(* IEC 61131-3 sources: Lasal-MCP/examples/SampleSource/5_ClassInputOutputSolution/Stations/MachineControl/MachineControl/Class/OPModeConfigBase, 1 file *)

(* ---- OPModeConfigBase.st ---- *)
#define     NewInstCmd_GetAlarms                  100     // newinst command to get alarms of station (class AlarmSation + class OPModeComMaster)
// parameter 1: sAlarmList  : t_s_OPMode
// parameter 2: bdAlarmInfo : BDINT

(*!
<Class
	Name               = "OPModeConfigBase"
	Revision           = "1.3"
	RealtimeTask       = "false"
	CyclicTask         = "false"
	BackgroundTask     = "false"
	Sigmatek           = "true"
	OSInterface        = "false"
	HighPriority       = "false"
	Automatic          = "false"
	UpdateMode         = "Prescan"
	SharedCommandTable = "true"
	Objectsize         = "(410,120)"
	Comment            = "This class defines the configuration for the class OPModeBase.&#13;&#10;All the possible ways to change the operation mode are defined within this class.&#13;&#10;&#13;&#10;Derive this class to change the configuration for switching the operation modes.">
	<Channels>
		<Server Name="ClassSvr" Visualized="false" Initialize="false" WriteProtected="true" Retentive="false"/>
	</Channels>
	<RevDoku>
		<Owner Company="Sigmatek" Author="ObeChr"/>
		<Dokumentation Revision="1.3" Date="2018-04-17" Author="ObeChr" Company="Sigmatek" Description="Added functionality that it is possible to call Change-Methods until every Slave Object is READY"/>
		<Dokumentation Revision="1.2" Date="2017-01-30" Author="ObeChr" Company="Sigmatek" Description="Added new public types to class."/>
		<Dokumentation Revision="1.1" Date="2016-03-08" Author="ObeChr" Company="Sigmatek" Description="+) Added deactivated configurations to the methods GetChangeConfig(), GetModeConfig() to show the possibilties of the class.&#13;&#10;+) Deactivated all transition times.&#13;&#10;+) Improved comments of global methods and variables."/>
		<Dokumentation Revision="1.0" Date="2015-06-01" Author="ObeChr" Company="Sigmatek" Description="First Version of class for the configuration of the operationmodes."/>
	</RevDoku>
</Class>
*)
OPModeConfigBase : CLASS
	TYPE
	  t_bd_OPMode : BDINT  //! <Type Public="true" Name="t_bd_OPMode"/>
	  [
	    1 bOPModeInit,
	    2 bOPModeHoming,
	    3 bOPModeStop,
	    4 bOPModeSetup,
	    5 bOPModeManual,
	    6 bOPModeSemiAuto,
	    7 bOPModeAutomatic,
	    8 bOPModeError,
	  ];
#pragma pack(push, 1)
	  t_s_OPChange : STRUCT  //! <Type Public="true" Name="t_s_OPChange"/>
	    bOPModeInit : BINT  //! <Type Comment="This bit field defines the optional operating modes to which are changed from the operating mode Init." Name="t_s_OPChange.bOPModeInit"/>
	    [
	      1 bHoming,
	      2 bStop,
	      3 bSetup,
	      4 bManual,
	      5 bSemiAuto,
	      6 bAutomatic,
	      7 bError,
	    ];
	    bOPModeHoming : BINT  //! <Type Comment="This bit field defines the optional operating modes to which are changed from the operating mode Homing." Name="t_s_OPChange.bOPModeHoming"/>
	    [
	      1 bInit,
	      2 bStop,
	      3 bSetup,
	      4 bManual,
	      5 bSemiAuto,
	      6 bAutomatic,
	      7 bError,
	    ];
	    bOPModeStop : BINT  //! <Type Comment="This bit field defines the optional operating modes to which are changed from the operating mode Stop." Name="t_s_OPChange.bOPModeStop"/>
	    [
	      1 bInit,
	      2 bHoming,
	      3 bSetup,
	      4 bManual,
	      5 bSemiAuto,
	      6 bAutomatic,
	      7 bError,
	    ];
	    bOPModeSetup : BINT  //! <Type Comment="This bit field defines the optional operating modes to which are changed from the operating mode Setup." Name="t_s_OPChange.bOPModeSetup"/>
	    [
	      1 bInit,
	      2 bHoming,
	      3 bStop,
	      4 bManual,
	      5 bSemiAuto,
	      6 bAutomatic,
	      7 bError,
	    ];
	    bOPModeManual : BINT  //! <Type Comment="This bit field defines the optional operating modes to which are changed from the operating mode Manual." Name="t_s_OPChange.bOPModeManual"/>
	    [
	      1 bInit,
	      2 bHoming,
	      3 bStop,
	      4 bSetup,
	      5 bSemiAuto,
	      6 bAutomatic,
	      7 bError,
	    ];
	    bOPModeSemiAuto : BINT  //! <Type Comment="This bit field defines the optional operating modes to which are changed from the operating mode SemiAuto." Name="t_s_OPChange.bOPModeSemiAuto"/>
	    [
	      1 bInit,
	      2 bHoming,
	      3 bStop,
	      4 bSetup,
	      5 bManual,
	      6 bAutomatic,
	      7 bError,
	    ];
	    bOPModeAutomatic : BINT  //! <Type Comment="This bit field defines the optional operating modes to which are changed from the operating mode Automatic." Name="t_s_OPChange.bOPModeAutomatic"/>
	    [
	      1 bInit,
	      2 bHoming,
	      3 bStop,
	      4 bSetup,
	      5 bManual,
	      6 bSemiAuto,
	      7 bError,
	    ];
	    bOPModeError : BINT  //! <Type Comment="This bit field defines the optional operating modes to which are changed from the operating mode Error." Name="t_s_OPChange.bOPModeError"/>
	    [
	      1 bInit,
	      2 bHoming,
	      3 bStop,
	      4 bSetup,
	      5 bManual,
	      6 bSemiAuto,
	      7 bAutomatic,
	    ];
	  END_STRUCT;
#pragma pack(pop)
#pragma pack(push, 1)
	  t_s_OPChangeTime : STRUCT  //! <Type Public="true" Name="t_s_OPChangeTime"/>
	    sOPModeInit : STRUCT  //! <Type Comment="In this structure, the allowable changeover times [ms] are defined from OPMode_Init.&#13;&#10;" Name="t_s_OPChangeTime.sOPModeInit"/>
	      udChangeToHoming : UDINT;
	      udChangeToStop : UDINT;
	      udChangeToSetup : UDINT;
	      udChangeToManual : UDINT;
	      udChangeToSemiAuto : UDINT;
	      udChangeToAutomatic : UDINT;
	      udChangeToError : UDINT;
	    END_STRUCT;
	    sOPModeHoming : STRUCT  //! <Type Comment="In this structure, the allowable changeover times [ms] are defined from OPMode_Homing.&#13;&#10;" Name="t_s_OPChangeTime.sOPModeHoming"/>
	      udChangeToInit : UDINT;
	      udChangeToStop : UDINT;
	      udChangeToSetup : UDINT;
	      udChangeToManual : UDINT;
	      udChangeToSemiAuto : UDINT;
	      udChangeToAutomatic : UDINT;
	      udChangeToError : UDINT;
	    END_STRUCT;
	    sOPModeStop : STRUCT  //! <Type Comment="In this structure, the allowable changeover times [ms] are defined from OPMode_Stop.&#13;&#10;" Name="t_s_OPChangeTime.sOPModeStop"/>
	      udChangeToInit : UDINT;
	      udChangeToHoming : UDINT;
	      udChangeToSetup : UDINT;
	      udChangeToManual : UDINT;
	      udChangeToSemiAuto : UDINT;
	      udChangeToAutomatic : UDINT;
	      udChangeToError : UDINT;
	    END_STRUCT;
	    sOPModeSetup : STRUCT  //! <Type Comment="In this structure, the allowable changeover times [ms] are defined from OPMode_Setup.&#13;&#10;" Name="t_s_OPChangeTime.sOPModeSetup"/>
	      udChangeToInit : UDINT;
	      udChangeToHoming : UDINT;
	      udChangeToStop : UDINT;
	      udChangeToManual : UDINT;
	      udChangeToSemiAuto : UDINT;
	      udChangeToAutomatic : UDINT;
	      udChangeToError : UDINT;
	    END_STRUCT;
	    sOPModeManual : STRUCT  //! <Type Comment="In this structure, the allowable changeover times [ms] are defined from OPMode_Manual.&#13;&#10;" Name="t_s_OPChangeTime.sOPModeManual"/>
	      udChangeToInit : UDINT;
	      udChangeToHoming : UDINT;
	      udChangeToStop : UDINT;
	      udChangeToSetup : UDINT;
	      udChangeToSemiAuto : UDINT;
	      udChangeToAutomatic : UDINT;
	      udChangeToError : UDINT;
	    END_STRUCT;
	    sOPModeSemiAuto : STRUCT  //! <Type Comment="In this structure, the allowable changeover times [ms] are defined from OPMode_SemiAuto.&#13;&#10;" Name="t_s_OPChangeTime.sOPModeSemiAuto"/>
	      udChangeToInit : UDINT;
	      udChangeToHoming : UDINT;
	      udChangeToStop : UDINT;
	      udChangeToSetup : UDINT;
	      udChangeToManual : UDINT;
	      udChangeToAutomatic : UDINT;
	      udChangeToError : UDINT;
	    END_STRUCT;
	    sOPModeAutomatic : STRUCT  //! <Type Comment="In this structure, the allowable changeover times [ms] are defined from OPMode_Automatic.&#13;&#10;" Name="t_s_OPChangeTime.sOPModeAutomatic"/>
	      udChangeToInit : UDINT;
	      udChangeToHoming : UDINT;
	      udChangeToStop : UDINT;
	      udChangeToSetup : UDINT;
	      udChangeToManual : UDINT;
	      udChangeToSemiAuto : UDINT;
	      udChangeToError : UDINT;
	    END_STRUCT;
	    sOPModeError : STRUCT  //! <Type Comment="In this structure, the allowable changeover times [ms] are defined from OPMode_Error.&#13;&#10;" Name="t_s_OPChangeTime.sOPModeError"/>
	      udChangeToInit : UDINT;
	      udChangeToHoming : UDINT;
	      udChangeToStop : UDINT;
	      udChangeToSetup : UDINT;
	      udChangeToManual : UDINT;
	      udChangeToSemiAuto : UDINT;
	      udChangeToAutomatic : UDINT;
	    END_STRUCT;
	  END_STRUCT;
#pragma pack(pop)
	END_TYPE
  //Servers:
	ClassSvr 	: SvrChCmd_DINT;
  //Clients:
  //Variables:
		bdOPMode 	: t_bd_OPMode;			//! <Variable Comment="This variable defines the available operation modes." Name="bdOPMode"/>
		sOPChange 	: t_s_OPChange;			//! <Variable Comment="This variable defines the possible transitions between the operation modes." Name="sOPChange"/>
		sOPChangeTime 	: t_s_OPChangeTime;			//! <Variable Comment="This variable defines the timeouts for the transitions between the operation modes." Name="sOPChangeTime"/>
  //Functions:
				//! <Function Comment="This method is called by the &quot;OPModeBase&quot; class during the last Init cycle. The configuration of the class is thereby defined. By overwriting this method, the default configuration can be changed." Name="GetChangeConfig"/>
	FUNCTION VIRTUAL GLOBAL GetChangeConfig
		VAR_OUTPUT
			pConfig 	: ^t_s_OPChange;			//! <Variable Comment="Pointer to the changeover options of the operating mode (sOPModeChange variable)." Name="GetChangeConfig.pConfig"/>
		END_VAR;
				//! <Function Comment="This method is called by the &quot;OPModeBase&quot; class during the last Init cycle. Through this call, the configuration is read based on allowed changeover time of the operating modes. By overwriting this method, the default configuration can be changed." Name="GetChangeTime"/>
	FUNCTION VIRTUAL GLOBAL GetChangeTime
		VAR_OUTPUT
			pConfig 	: ^t_s_OPChangeTime;			//! <Variable Comment="Pointer to the timeouts when changing operating modes  (variable sOPChangeTime)." Name="GetChangeTime.pConfig"/>
		END_VAR;
				//! <Function Comment="This method is called by the &quot;AlarmBufferBase&quot; class when registering an alarm. The possible configuration of the alarm is checked. By overwriting this method, the default configuration can be changed." Name="GetModeConfig"/>
	FUNCTION VIRTUAL GLOBAL GetModeConfig
		VAR_OUTPUT
			pConfig 	: ^t_bd_OPMode;			//! <Variable Comment="Pointer to the available operating modes (variable bdOPMode)." Name="GetModeConfig.pConfig"/>
		END_VAR;
  //Tables:
	FUNCTION @STD
		VAR_OUTPUT
			ret_code	: CONFSTATES;
		END_VAR;
	FUNCTION GLOBAL TAB @CT_;
END_CLASS;

FUNCTION VIRTUAL GLOBAL OPModeConfigBase::GetChangeConfig
	VAR_OUTPUT
		pConfig 	: ^t_s_OPChange;
	END_VAR

  // this information is ued by the class OPModeBase
  // => only following transitions between the OPModes
  //    can be used

  // possibilities to leave OPMode_Init
  sOPChange.bOPModeInit.bHoming     := true;        // transition active
  sOPChange.bOPModeInit.bStop       := false;
  sOPChange.bOPModeInit.bSetup      := false;
  sOPChange.bOPModeInit.bManual     := false;
  sOPChange.bOPModeInit.bSemiAuto   := false;
  sOPChange.bOPModeInit.bAutomatic  := false;
  sOPChange.bOPModeInit.bError      := true;        // transition active

  // possibilities to leave OPMode_Homing
  sOPChange.bOPModeHoming.bInit       := false;
  sOPChange.bOPModeHoming.bStop       := false;
  sOPChange.bOPModeHoming.bSetup      := false;
  sOPChange.bOPModeHoming.bManual     := true;      // transition active
  sOPChange.bOPModeHoming.bSemiAuto   := false;
  sOPChange.bOPModeHoming.bAutomatic  := false;
  sOPChange.bOPModeHoming.bError      := true;      // transition active

  // possibilities to leave OPMode_Stop
  sOPChange.bOPModeStop.bInit       := false;
  sOPChange.bOPModeStop.bHoming     := false;
  sOPChange.bOPModeStop.bSetup      := false;
  sOPChange.bOPModeStop.bManual     := false;
  sOPChange.bOPModeStop.bSemiAuto   := false;
  sOPChange.bOPModeStop.bAutomatic  := false;
  sOPChange.bOPModeStop.bError      := false;

  // possibilities to leave OPMode_Setup
  sOPChange.bOPModeSetup.bInit      := false;
  sOPChange.bOPModeSetup.bHoming    := false;
  sOPChange.bOPModeSetup.bStop      := false;
  sOPChange.bOPModeSetup.bManual    := false;
  sOPChange.bOPModeSetup.bSemiAuto  := false;
  sOPChange.bOPModeSetup.bAutomatic := false;
  sOPChange.bOPModeSetup.bError     := false;

  // possibilities to leave OPMode_Manual
  sOPChange.bOPModeManual.bInit       := true;      // transition active
  sOPChange.bOPModeManual.bHoming     := true;      // transition active
  sOPChange.bOPModeManual.bStop       := false;
  sOPChange.bOPModeManual.bSetup      := false;
  sOPChange.bOPModeManual.bSemiAuto   := true;      // transition active
  sOPChange.bOPModeManual.bAutomatic  := true;      // transition active
  sOPChange.bOPModeManual.bError      := true;      // transition active

  // possibilities to leave OPMode_SemiAuto
  sOPChange.bOPModeSemiAuto.bInit       := false;
  sOPChange.bOPModeSemiAuto.bHoming     := false;
  sOPChange.bOPModeSemiAuto.bStop       := false;
  sOPChange.bOPModeSemiAuto.bSetup      := false;
  sOPChange.bOPModeSemiAuto.bManual     := true;    // transition active
  sOPChange.bOPModeSemiAuto.bAutomatic  := true;    // transition active
  sOPChange.bOPModeSemiAuto.bError      := true;    // transition active

  // possibilities to leave OPMode_Automatic
  sOPChange.bOPModeAutomatic.bInit      := false;
  sOPChange.bOPModeAutomatic.bHoming    := false;
  sOPChange.bOPModeAutomatic.bStop      := false;
  sOPChange.bOPModeAutomatic.bSetup     := false;
  sOPChange.bOPModeAutomatic.bManual    := true;    // transition active
  sOPChange.bOPModeAutomatic.bSemiAuto  := true;    // transition active
  sOPChange.bOPModeAutomatic.bError     := true;    // transition active

  // possibilities to leave OPMode_Error
  sOPChange.bOPModeError.bInit      := true;        // transition active
  sOPChange.bOPModeError.bHoming    := true;        // transition active
  sOPChange.bOPModeError.bStop      := false;
  sOPChange.bOPModeError.bSetup     := false;
  sOPChange.bOPModeError.bManual    := true;        // transition active
  sOPChange.bOPModeError.bSemiAuto  := false;
  sOPChange.bOPModeError.bAutomatic := false;

  // return pointer to configuration
  pConfig := #sOPChange;

END_FUNCTION

FUNCTION VIRTUAL GLOBAL OPModeConfigBase::GetModeConfig
	VAR_OUTPUT
		pConfig 	: ^t_bd_OPMode;
	END_VAR

  // this information is used by the class AlarmBuffer
  // => only following OPModes can be set at the alarm
  //    objects

  // available OPModes
  bdOPMode.bOPModeInit      := true;    // OPMode active
  bdOPMode.bOPModeHoming    := true;    // OPMode active
  bdOPMode.bOPModeStop      := false;
  bdOPMode.bOPModeSetup     := false;
  bdOPMode.bOPModeManual    := true;    // OPMode active
  bdOPMode.bOPModeSemiAuto  := true;    // OPMode active
  bdOPMode.bOPModeAutomatic := true;    // OPMode active
  bdOPMode.bOPModeError     := true;    // OPMode active

  // return configuration
  pConfig := #bdOPMode;

END_FUNCTION

FUNCTION VIRTUAL GLOBAL OPModeConfigBase::GetChangeTime
	VAR_OUTPUT
		pConfig 	: ^t_s_OPChangeTime;
	END_VAR

  // this information is ued by the class OPModeBase
  // => in case changing the opmode takes more than
  //    the selected time, an error occus.
  // 0: check of transitiontime is deactivated

  // timeouts to leave OPMode_Init
  sOPChangeTime.sOPModeInit.udChangeToHoming    := 0;
  sOPChangeTime.sOPModeInit.udChangeToStop      := 0;
  sOPChangeTime.sOPModeInit.udChangeToSetup     := 0;
  sOPChangeTime.sOPModeInit.udChangeToManual    := 0;
  sOPChangeTime.sOPModeInit.udChangeToSemiAuto  := 0;
  sOPChangeTime.sOPModeInit.udChangeToAutomatic := 0;
  sOPChangeTime.sOPModeInit.udChangeToError     := 0;

  // timeouts to leave OPMode_Homing
  sOPChangeTime.sOPModeHoming.udChangeToInit      := 0;
  sOPChangeTime.sOPModeHoming.udChangeToStop      := 0;
  sOPChangeTime.sOPModeHoming.udChangeToSetup     := 0;
  sOPChangeTime.sOPModeHoming.udChangeToManual    := 0;
  sOPChangeTime.sOPModeHoming.udChangeToSemiAuto  := 0;
  sOPChangeTime.sOPModeHoming.udChangeToAutomatic := 0;
  sOPChangeTime.sOPModeHoming.udChangeToError     := 0;

  // timeouts to leave OPMode_Stop
  sOPChangeTime.sOPModeStop.udChangeToInit      := 0;
  sOPChangeTime.sOPModeStop.udChangeToHoming    := 0;
  sOPChangeTime.sOPModeStop.udChangeToSetup     := 0;
  sOPChangeTime.sOPModeStop.udChangeToManual    := 0;
  sOPChangeTime.sOPModeStop.udChangeToSemiAuto  := 0;
  sOPChangeTime.sOPModeStop.udChangeToAutomatic := 0;
  sOPChangeTime.sOPModeStop.udChangeToError     := 0;

  // timeouts to leave OPMode_Setup
  sOPChangeTime.sOPModeSetup.udChangeToInit       := 0;
  sOPChangeTime.sOPModeSetup.udChangeToHoming     := 0;
  sOPChangeTime.sOPModeSetup.udChangeToStop       := 0;
  sOPChangeTime.sOPModeSetup.udChangeToManual     := 0;
  sOPChangeTime.sOPModeSetup.udChangeToSemiAuto   := 0;
  sOPChangeTime.sOPModeSetup.udChangeToAutomatic  := 0;
  sOPChangeTime.sOPModeSetup.udChangeToError      := 0;

  // timeouts to leave OPMode_Manual
  sOPChangeTime.sOPModeManual.udChangeToInit      := 0;
  sOPChangeTime.sOPModeManual.udChangeToHoming    := 0;
  sOPChangeTime.sOPModeManual.udChangeToStop      := 0;
  sOPChangeTime.sOPModeManual.udChangeToSetup     := 0;
  sOPChangeTime.sOPModeManual.udChangeToSemiAuto  := 0;
  sOPChangeTime.sOPModeManual.udChangeToAutomatic := 0;
  sOPChangeTime.sOPModeManual.udChangeToError     := 0;

  // timeouts to leave OPMode_SemiAuto
  sOPChangeTime.sOPModeSemiAuto.udChangeToInit      := 0;
  sOPChangeTime.sOPModeSemiAuto.udChangeToHoming    := 0;
  sOPChangeTime.sOPModeSemiAuto.udChangeToStop      := 0;
  sOPChangeTime.sOPModeSemiAuto.udChangeToSetup     := 0;
  sOPChangeTime.sOPModeSemiAuto.udChangeToManual    := 0;
  sOPChangeTime.sOPModeSemiAuto.udChangeToAutomatic := 0;
  sOPChangeTime.sOPModeSemiAuto.udChangeToError     := 0;

  // timeouts to leave OPMode_Automatic
  sOPChangeTime.sOPModeAutomatic.udChangeToInit     := 0;
  sOPChangeTime.sOPModeAutomatic.udChangeToHoming   := 0;
  sOPChangeTime.sOPModeAutomatic.udChangeToStop     := 0;
  sOPChangeTime.sOPModeAutomatic.udChangeToSetup    := 0;
  sOPChangeTime.sOPModeAutomatic.udChangeToManual   := 0;
  sOPChangeTime.sOPModeAutomatic.udChangeToSemiAuto := 0;
  sOPChangeTime.sOPModeAutomatic.udChangeToError    := 0;

  // timeouts to leave OPMode_Error
  sOPChangeTime.sOPModeError.udChangeToInit       := 0;
  sOPChangeTime.sOPModeError.udChangeToHoming     := 0;
  sOPChangeTime.sOPModeError.udChangeToStop       := 0;
  sOPChangeTime.sOPModeError.udChangeToSetup      := 0;
  sOPChangeTime.sOPModeError.udChangeToManual     := 0;
  sOPChangeTime.sOPModeError.udChangeToSemiAuto   := 0;
  sOPChangeTime.sOPModeError.udChangeToAutomatic  := 0;

  // return pointer to configuration
  pConfig := #sOPChangeTime;

END_FUNCTION
